TYPE ST_GFX4IR_REF : FB_GFX4IR_REF;
END_TYPE

(* stored: Version 1.1.0.1, ProductVersion 3.1.4024.15
   DUT ST_GFX4IR_REF: Id {fbefe143-8609-4a6d-9fdb-fe06f5882f36} *)
